// SIMATIC S7-200 project (STEP 7-Micro/WIN), CPU 226 CN REL 02.01

SYMBOL_TABLE Tabla de símbolos
QS               I2.6     // BOTON DE EMERGENCIA
SB_1             I2.5     // PULSADOR DE MARCHA
SB_2             I2.4     // PULSADOR DE PARO
SA               I2.7     // SELECTOR
SPSS             I0.7     // SENSOR PISTON SUJETADOR SALE
SPLE             I0.6     // SENSOR PISTON LIBERADOR ENRA
SPLS             I0.5     // SENSOR PISTON LIBERADOR SALE
SPSE             I1.0     // SENSOR PISTON SUJETADOR ENTRA
SST              I0.2     // SENSOR SALIDA TUBO
SGA              I1.1     // SENSOR GIRO ANTI-HORAIO
SPR              I0.3     // SENSOR PRESENFCIA RECOGER
SGRA             I1.3     // SENSOR GARRA ABIERTO
SFO              I0.4     // SENSOR DEPOSITO
SGRS             I1.5     // SENSOR GARRA SUBE
SGH              I1.2     // SENSOR GIRO HORARIO
SGRB             I1.4     // SENSOR GARRA BAJA
SGRAD            I1.7     // SENSOR GARRA ADELANTE
SGRT             I1.6     // SENSOR GARRA HORIZONTAL ATRAS
ST_I             I0.0     // SENSOR TUBO INFERIOR
PLIB             Q0.1     // PISTON LIBERADOR
PSUJ             Q0.0     // PISTON SUJETADOR
CILROTAH         Q0.2     // CILINDRO ROTATORIO ANTI-HORARIO
CILHORADE        Q0.5     // CILINDRO HORIZONTAL ADELANTE
CILVERTABAJO     Q0.4     // CILINDRO VERTICAL ABAJO
FINGER           Q0.3     // GARRA CIERRA
HA               Q1.5     // LAMPARA AMARILLA
HV               Q1.6     // LAMPARA VERDE
HR               Q1.7     // LAMPARA ROJA
BALY             Q0.7     // BALIZA AMARILLO
BALV             Q1.0     // BALIZA VERDE
E0               M0.0
E1               M0.1
E2               M0.2
E3               M0.3
E4               M0.4
E5               M0.5
E6               M0.6
E7               M0.7
E8               M1.0
E9               M1.1
E10              M1.2
E11              M1.3
E12              M1.4
E13              M1.5
E14              M1.6
E15              M2.1
E16              M1.7     // ESTADO DE EMERGENCIA
STOPP            M2.0     // PARADA MOMENTANEA
COM_FINALIZADO   V0.3
COM_INICIAR      V0.2
END_SYMBOL_TABLE

ORGANIZATION_BLOCK Bloque_de_programa:OB1
TITLE=COMENTARIOS DEL PROGRAMA
BEGIN
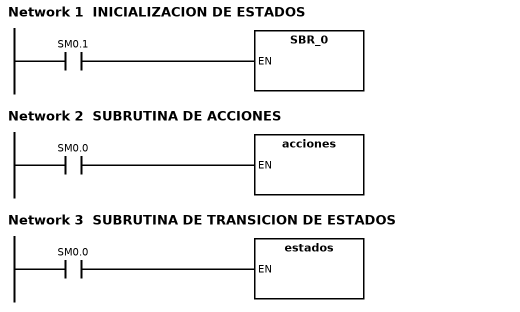
Network 1 // INICIALIZACION DE ESTADOS
LD     SM0.1
CALL   SBR_0:SBR0
Network 2 // SUBRUTINA DE ACCIONES
LD     SM0.0
CALL   acciones:SBR1
Network 3 // SUBRUTINA DE TRANSICION DE ESTADOS
LD     SM0.0
CALL   estados:SBR2
END_ORGANIZATION_BLOCK

SUBROUTINE_BLOCK SBR_0:SBR0
TITLE=COMENTARIOS DE LA SUBRUTINA
BEGIN
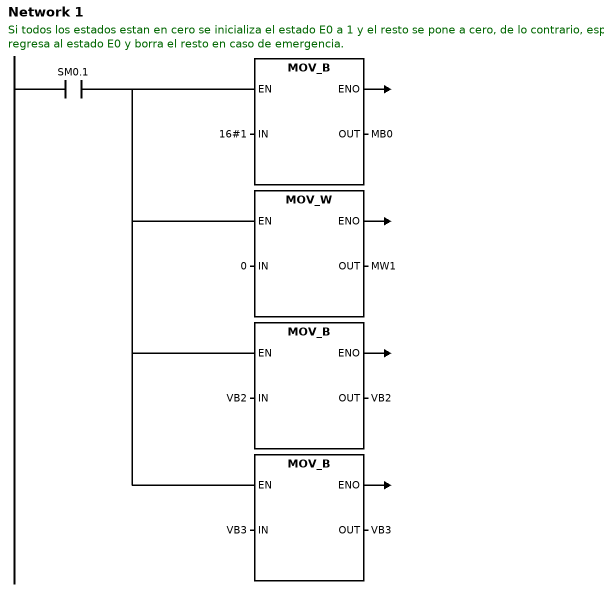
Network 1
// Si todos los estados estan en cero se inicializa el estado E0 a 1 y el resto se pone a cero, de lo contrario, espera a que se oprima el boton de emergencia. Tambien es la manera en que el programa regresa al estado E0 y borra el resto en caso de emergencia.
LD     SM0.1
MOVB   16#1, MB0
MOVW   0, MW1
MOVB   VB2, VB2
MOVB   VB3, VB3
END_SUBROUTINE_BLOCK

SUBROUTINE_BLOCK acciones:SBR1
TITLE=COMENTARIOS DE LA SUBRUTINA
BEGIN
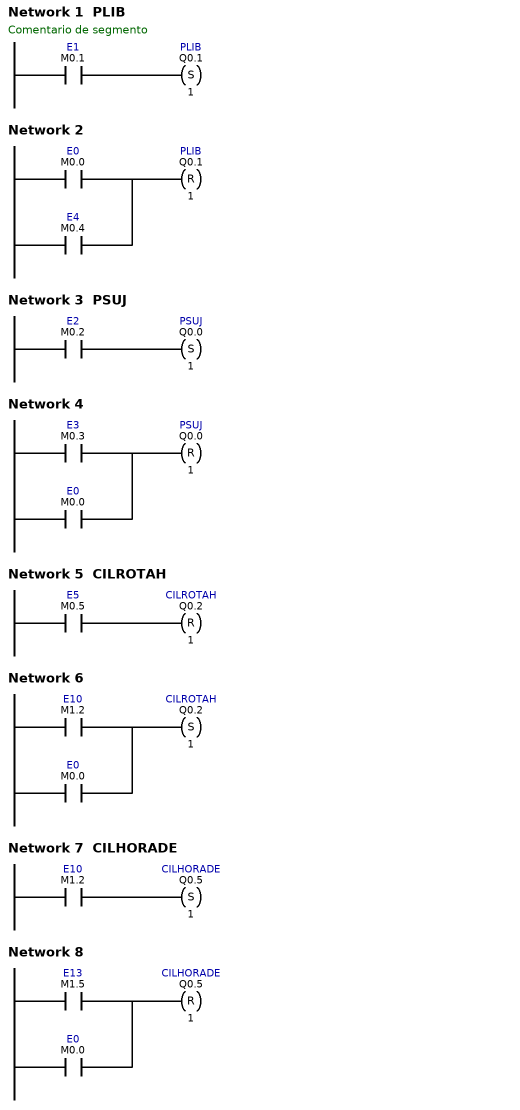
Network 1 // PLIB
// Comentario de segmento
LD     E1:M0.1
S      PLIB:Q0.1, 1
Network 2
LD     E0:M0.0
O      E4:M0.4
R      PLIB:Q0.1, 1
Network 3 // PSUJ
LD     E2:M0.2
S      PSUJ:Q0.0, 1
Network 4
LD     E3:M0.3
O      E0:M0.0
R      PSUJ:Q0.0, 1
Network 5 // CILROTAH
LD     E5:M0.5
R      CILROTAH:Q0.2, 1
Network 6
LD     E10:M1.2
O      E0:M0.0
S      CILROTAH:Q0.2, 1
Network 7 // CILHORADE
LD     E10:M1.2
S      CILHORADE:Q0.5, 1
Network 8
LD     E13:M1.5
O      E0:M0.0
R      CILHORADE:Q0.5, 1
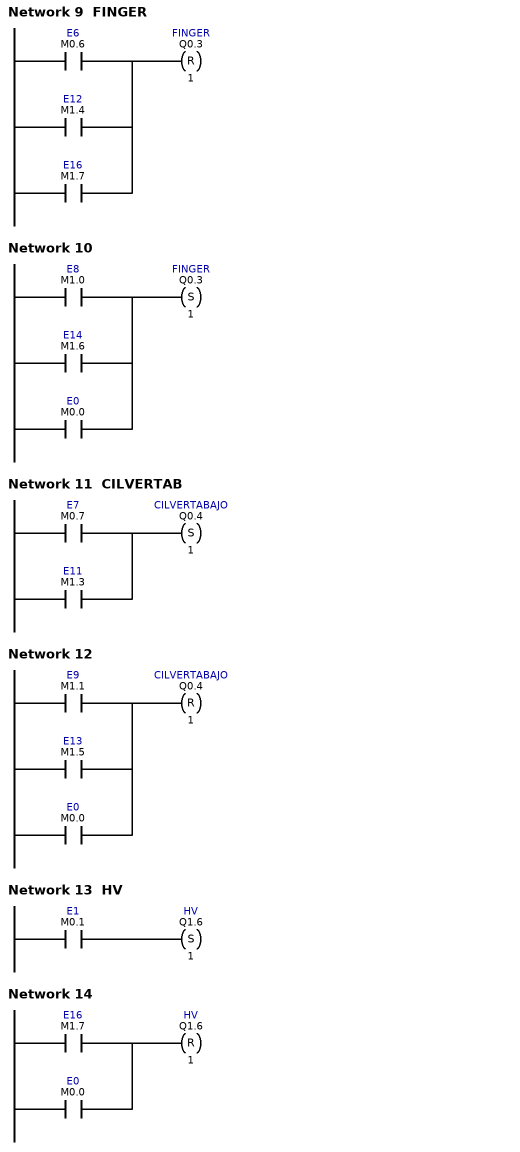
Network 9 // FINGER
LD     E6:M0.6
O      E12:M1.4
O      E16:M1.7
R      FINGER:Q0.3, 1
Network 10
LD     E8:M1.0
O      E14:M1.6
O      E0:M0.0
S      FINGER:Q0.3, 1
Network 11 // CILVERTAB
LD     E7:M0.7
O      E11:M1.3
S      CILVERTABAJO:Q0.4, 1
Network 12
LD     E9:M1.1
O      E13:M1.5
O      E0:M0.0
R      CILVERTABAJO:Q0.4, 1
Network 13 // HV
LD     E1:M0.1
S      HV:Q1.6, 1
Network 14
LD     E16:M1.7
O      E0:M0.0
R      HV:Q1.6, 1
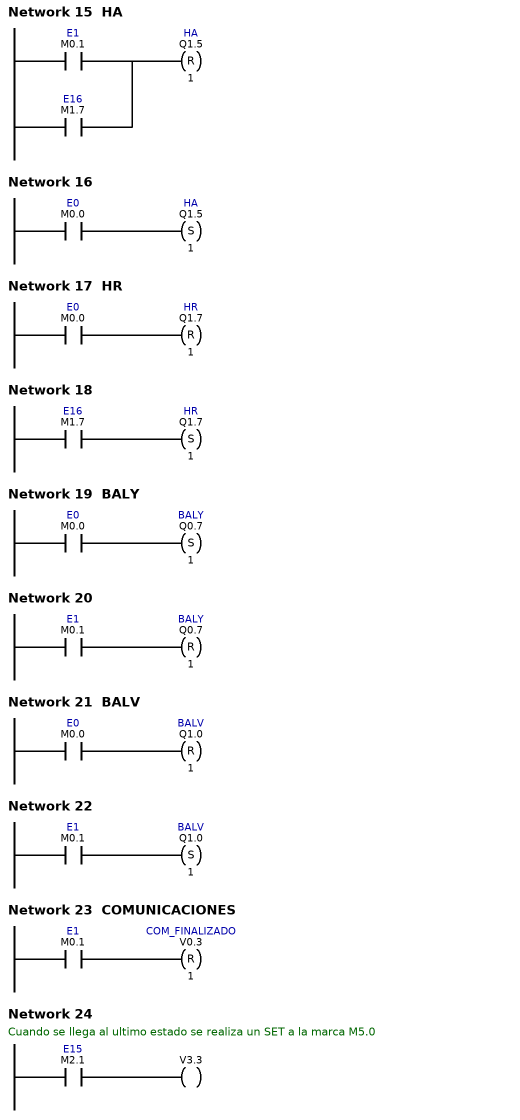
Network 15 // HA
LD     E1:M0.1
O      E16:M1.7
R      HA:Q1.5, 1
Network 16
LD     E0:M0.0
S      HA:Q1.5, 1
Network 17 // HR
LD     E0:M0.0
R      HR:Q1.7, 1
Network 18
LD     E16:M1.7
S      HR:Q1.7, 1
Network 19 // BALY
LD     E0:M0.0
S      BALY:Q0.7, 1
Network 20
LD     E1:M0.1
R      BALY:Q0.7, 1
Network 21 // BALV
LD     E0:M0.0
R      BALV:Q1.0, 1
Network 22
LD     E1:M0.1
S      BALV:Q1.0, 1
Network 23 // COMUNICACIONES
LD     E1:M0.1
R      COM_FINALIZADO:V0.3, 1
Network 24
// Cuando se llega al ultimo estado se realiza un SET a la marca M5.0
LD     E15:M2.1
=      V3.3
END_SUBROUTINE_BLOCK

SUBROUTINE_BLOCK estados:SBR2
TITLE=TRANSICION DE ESTADOS
BEGIN
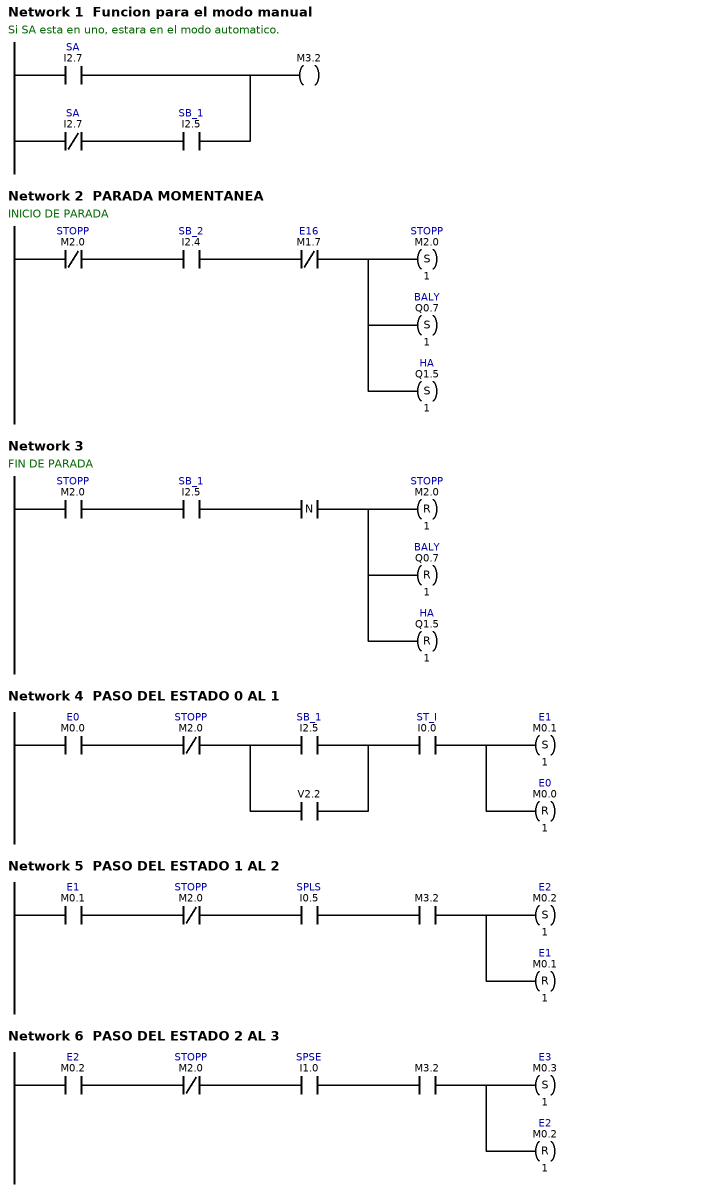
Network 1 // Funcion para el modo manual
// Si SA esta en uno, estara en el modo automatico. 
LD     SA:I2.7
LDN    SA:I2.7
A      SB_1:I2.5
OLD
=      M3.2
Network 2 // PARADA MOMENTANEA
// INICIO DE PARADA
LDN    STOPP:M2.0
A      SB_2:I2.4
AN     E16:M1.7
S      STOPP:M2.0, 1
S      BALY:Q0.7, 1
S      HA:Q1.5, 1
Network 3
// FIN DE PARADA
LD     STOPP:M2.0
A      SB_1:I2.5
ED
R      STOPP:M2.0, 1
R      BALY:Q0.7, 1
R      HA:Q1.5, 1
Network 4 // PASO DEL ESTADO 0 AL 1
LD     E0:M0.0
AN     STOPP:M2.0
LD     SB_1:I2.5
O      V2.2
ALD
A      ST_I:I0.0
S      E1:M0.1, 1
R      E0:M0.0, 1
Network 5 // PASO DEL ESTADO 1 AL 2
LD     E1:M0.1
AN     STOPP:M2.0
A      SPLS:I0.5
A      M3.2
S      E2:M0.2, 1
R      E1:M0.1, 1
Network 6 // PASO DEL ESTADO 2 AL 3
LD     E2:M0.2
AN     STOPP:M2.0
A      SPSE:I1.0
A      M3.2
S      E3:M0.3, 1
R      E2:M0.2, 1
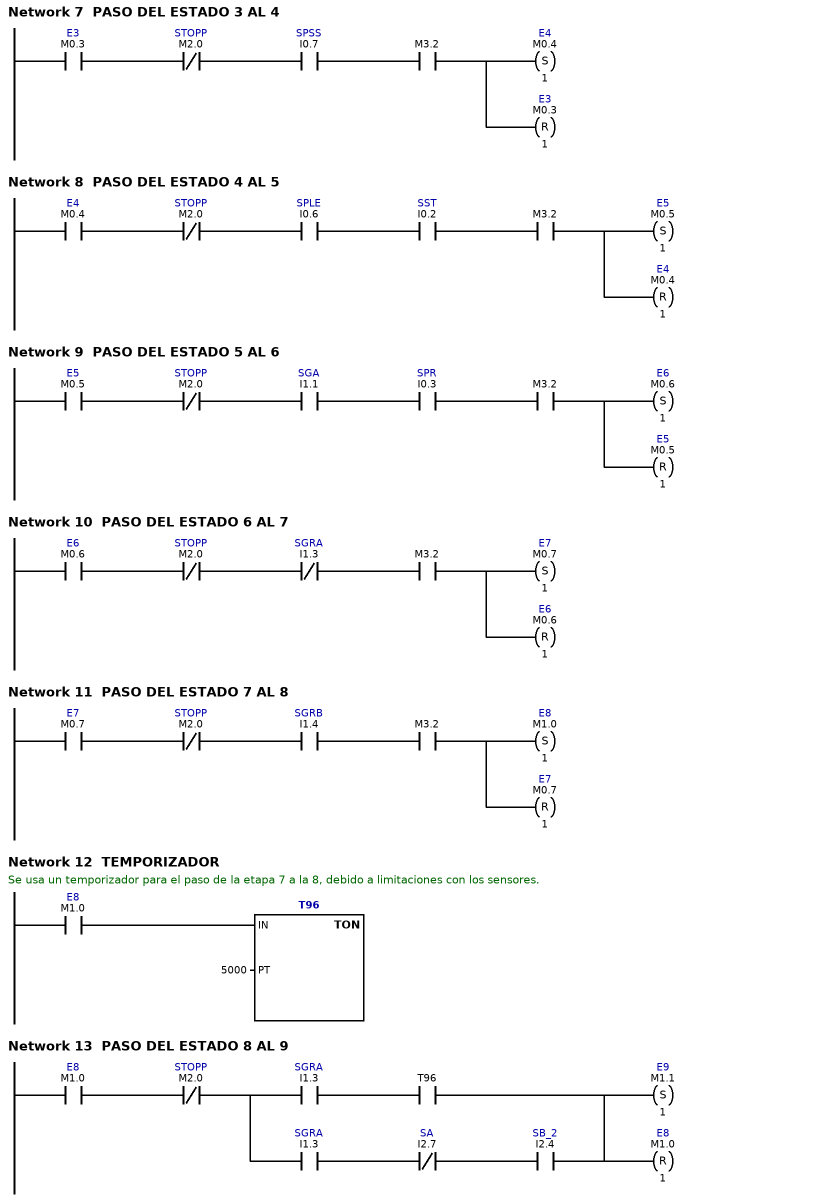
Network 7 // PASO DEL ESTADO 3 AL 4
LD     E3:M0.3
AN     STOPP:M2.0
A      SPSS:I0.7
A      M3.2
S      E4:M0.4, 1
R      E3:M0.3, 1
Network 8 // PASO DEL ESTADO 4 AL 5
LD     E4:M0.4
AN     STOPP:M2.0
A      SPLE:I0.6
A      SST:I0.2
A      M3.2
S      E5:M0.5, 1
R      E4:M0.4, 1
Network 9 // PASO DEL ESTADO 5 AL 6
LD     E5:M0.5
AN     STOPP:M2.0
A      SGA:I1.1
A      SPR:I0.3
A      M3.2
S      E6:M0.6, 1
R      E5:M0.5, 1
Network 10 // PASO DEL ESTADO 6 AL 7
LD     E6:M0.6
AN     STOPP:M2.0
AN     SGRA:I1.3
A      M3.2
S      E7:M0.7, 1
R      E6:M0.6, 1
Network 11 // PASO DEL ESTADO 7 AL 8
LD     E7:M0.7
AN     STOPP:M2.0
A      SGRB:I1.4
A      M3.2
S      E8:M1.0, 1
R      E7:M0.7, 1
Network 12 // TEMPORIZADOR
// Se usa un temporizador para el paso de la etapa 7 a la 8, debido a limitaciones con los sensores.
LD     E8:M1.0
TON    T96, 5000
Network 13 // PASO DEL ESTADO 8 AL 9
LD     E8:M1.0
AN     STOPP:M2.0
LD     SGRA:I1.3
A      T96
LD     SGRA:I1.3
AN     SA:I2.7
A      SB_2:I2.4
OLD
ALD
S      E9:M1.1, 1
R      E8:M1.0, 1
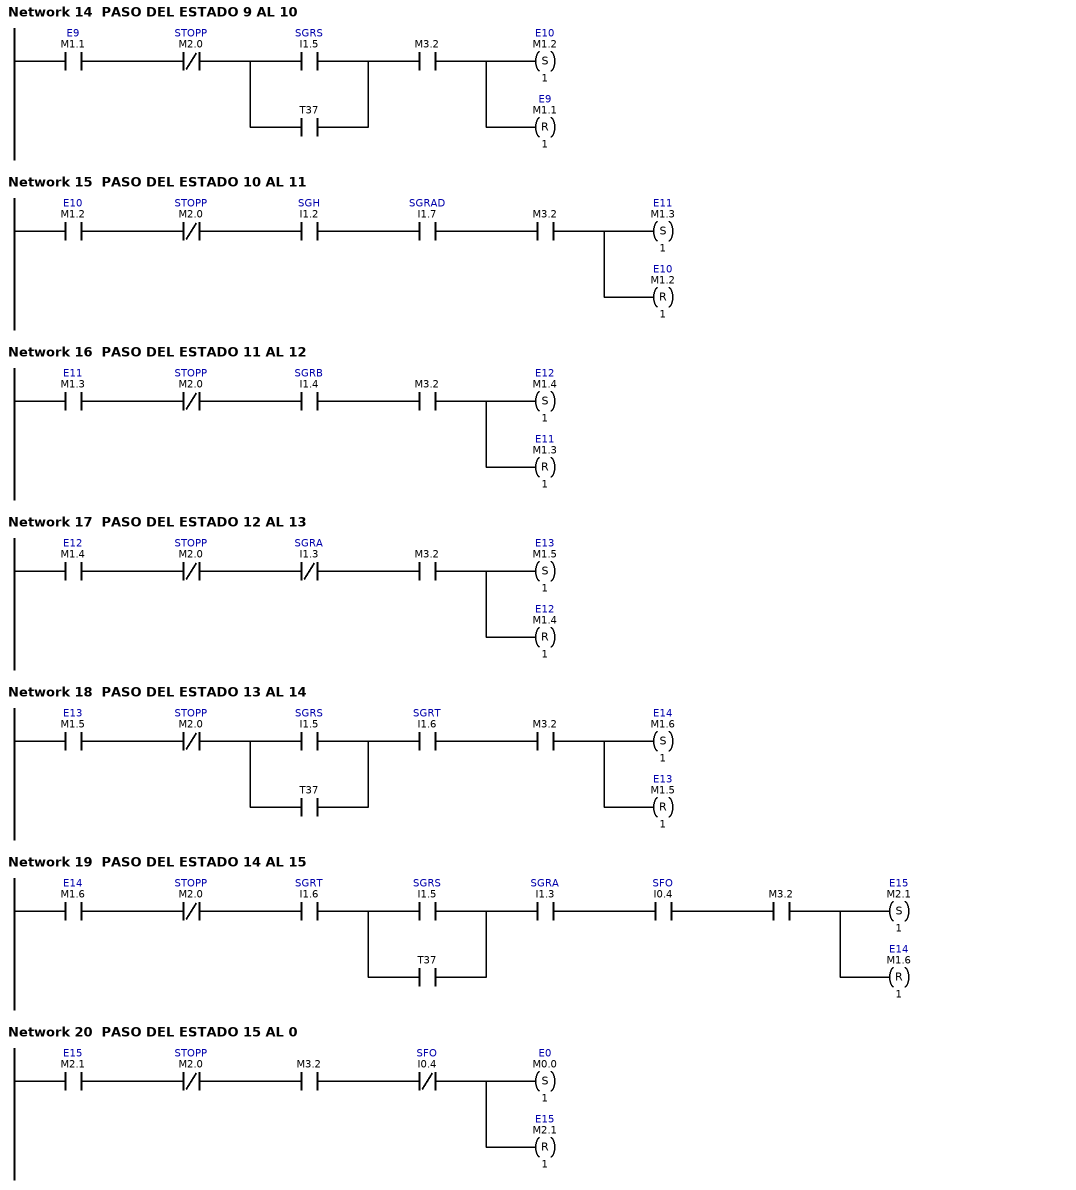
Network 14 // PASO DEL ESTADO 9 AL 10
LD     E9:M1.1
AN     STOPP:M2.0
LD     SGRS:I1.5
O      T37
ALD
A      M3.2
S      E10:M1.2, 1
R      E9:M1.1, 1
Network 15 // PASO DEL ESTADO 10 AL 11
LD     E10:M1.2
AN     STOPP:M2.0
A      SGH:I1.2
A      SGRAD:I1.7
A      M3.2
S      E11:M1.3, 1
R      E10:M1.2, 1
Network 16 // PASO DEL ESTADO 11 AL 12
LD     E11:M1.3
AN     STOPP:M2.0
A      SGRB:I1.4
A      M3.2
S      E12:M1.4, 1
R      E11:M1.3, 1
Network 17 // PASO DEL ESTADO 12 AL 13
LD     E12:M1.4
AN     STOPP:M2.0
AN     SGRA:I1.3
A      M3.2
S      E13:M1.5, 1
R      E12:M1.4, 1
Network 18 // PASO DEL ESTADO 13 AL 14
LD     E13:M1.5
AN     STOPP:M2.0
LD     SGRS:I1.5
O      T37
ALD
A      SGRT:I1.6
A      M3.2
S      E14:M1.6, 1
R      E13:M1.5, 1
Network 19 // PASO DEL ESTADO 14 AL 15
LD     E14:M1.6
AN     STOPP:M2.0
A      SGRT:I1.6
LD     SGRS:I1.5
O      T37
ALD
A      SGRA:I1.3
A      SFO:I0.4
A      M3.2
S      E15:M2.1, 1
R      E14:M1.6, 1
Network 20 // PASO DEL ESTADO 15 AL 0
LD     E15:M2.1
AN     STOPP:M2.0
A      M3.2
AN     SFO:I0.4
S      E0:M0.0, 1
R      E15:M2.1, 1
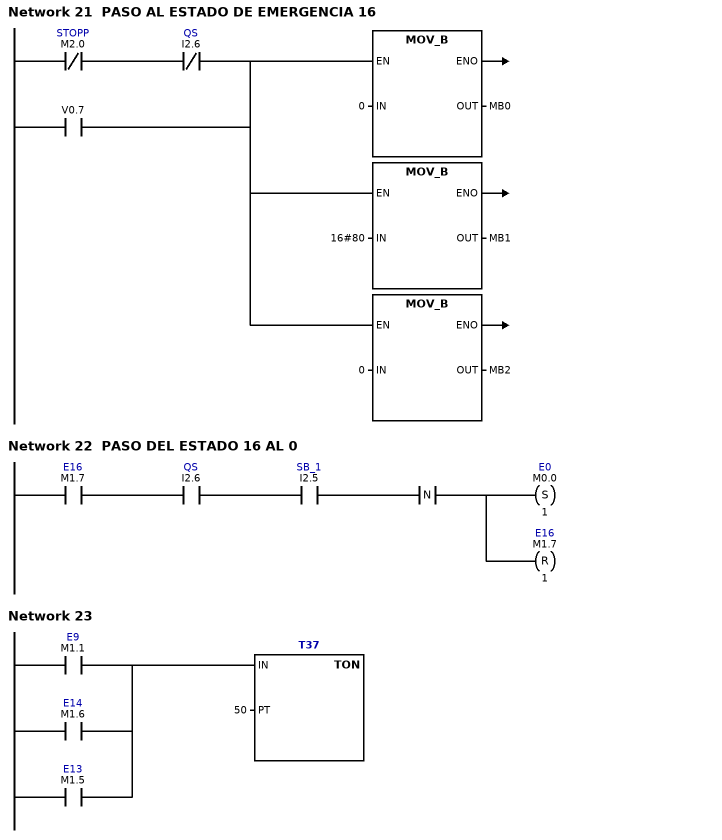
Network 21 // PASO AL ESTADO DE EMERGENCIA 16
LDN    STOPP:M2.0
AN     QS:I2.6
O      V0.7
MOVB   0, MB0
MOVB   16#80, MB1
MOVB   0, MB2
Network 22 // PASO DEL ESTADO 16 AL 0
LD     E16:M1.7
A      QS:I2.6
A      SB_1:I2.5
ED
S      E0:M0.0, 1
R      E16:M1.7, 1
Network 23
LD     E9:M1.1
O      E14:M1.6
O      E13:M1.5
TON    T37, 50
END_SUBROUTINE_BLOCK
